Fanuc KAREL source: kd00017.compact.KL

PROGRAM KD00017
%STACKSIZE=65535
%PRIORITY=65535
%NOLOCKGROUP
VAR
I : INTEGER
J : INTEGER
B : BOOLEAN
R : REAL
S : STRING[80]
BEGIN
I=0
CONNECT TIMER TO I
DISCONNECT TIMER I
END KD00017
